(* IEC 61131-3 sources: llm-plc-st-eval/data/processed_definitivo/qwen2.5-coder_14b/B7/zero_shot, 3 files *)

(* ---- ejec_1.st ---- *)
PROGRAM SelBomba
VAR
    modoAuto : BOOL;    // Entrada que indica el modo automático
    btnManual : BOOL;   // Entrada que indica el botón manual
    nivelBajo : BOOL;  // Entrada que indica el nivel bajo
    bomba : BOOL;       // Salida que indica el estado de la bomba
END_VAR

// Lógica de selección de la fuente de mando de la bomba
IF modoAuto THEN
    // Modo automático: la bomba está encendida si nivelBajo está activo
    bomba := nivelBajo;
ELSE
    // Modo manual: la bomba obedece al botón btnManual
    bomba := btnManual;
END_IF;

(* ---- ejec_2.st ---- *)
PROGRAM SelBomba
VAR
    modoAuto : BOOL;  // Entrada que indica si el sistema está en modo automático
    btnManual : BOOL; // Entrada que indica el estado del botón manual
    nivelBajo : BOOL; // Entrada que indica si el nivel está por debajo del umbral
    bomba : BOOL;     // Salida que indica el estado de la bomba
END_VAR

// Lógica de selección de la fuente de mando de la bomba
IF modoAuto THEN
    // En modo automático, la bomba está encendida si nivelBajo está activo
    bomba := nivelBajo;
ELSE
    // En modo manual, la bomba obedece directamente al botón btnManual
    bomba := btnManual;
END_IF;

(* ---- ejec_3.st ---- *)
PROGRAM SelBomba
VAR
    modoAuto : BOOL;   // Entrada que indica si el sistema está en modo automático
    btnManual : BOOL;  // Entrada que indica el estado del botón manual
    nivelBajo : BOOL;  // Entrada que indica si el nivel está por debajo del umbral
    bomba : BOOL;      // Salida que indica el estado de la bomba
END_VAR

// Lógica de selección de la fuente de mando de la bomba
IF modoAuto THEN
    // En modo automático, la bomba está encendida si nivelBajo está activo
    bomba := nivelBajo;
ELSE
    // En modo manual, la bomba obedece al botón manual
    bomba := btnManual;
END_IF;
